{attribute 'linkalways'}
{attribute 'no_explicit_call' := 'Use the methods of this class'}
{attribute 'enable_dynamic_creation'}
FUNCTION_BLOCK DiffDrive IMPLEMENTS I_DifferentialDrive
VAR
	leftAxis : I_DriveAxis;
	rightAxis : I_DriveAxis;
	kinematics : DiffDriveKinematics;
END_VAR

METHOD Connect
VAR_INPUT
	left : I_DriveAxis;
	right : I_DriveAxis;
END_VAR
leftAxis := left;
rightAxis := right;
END_METHOD

METHOD Execute
IF leftAxis = 0 OR rightAxis = 0 THEN
	RETURN;
END_IF
leftAxis.Execute();
rightAxis.Execute();
END_METHOD

METHOD Enable
IF leftAxis = 0 OR rightAxis = 0 THEN
	RETURN;
END_IF
leftAxis.Enable();
rightAxis.Enable();
END_METHOD

METHOD Disable
IF leftAxis = 0 OR rightAxis = 0 THEN
	RETURN;
END_IF
leftAxis.Disable();
rightAxis.Disable();
END_METHOD

METHOD SetTwist
VAR_INPUT
	desiredTwist : Twist;
END_VAR
VAR
	speeds : WheelSpeeds;
END_VAR
IF leftAxis = 0 OR rightAxis = 0 THEN
	RETURN;
END_IF
speeds := kinematics.ToWheelSpeeds(desiredTwist);
leftAxis.SetVelocity(speeds.leftInMPerS);
rightAxis.SetVelocity(speeds.rightInMPerS);
END_METHOD

PROPERTY LeftWheelPositionInM : LREAL
GET
IF leftAxis <> 0 THEN
	LeftWheelPositionInM := leftAxis.PositionInM;
END_IF
END_GET
END_PROPERTY

PROPERTY RightWheelPositionInM : LREAL
GET
IF rightAxis <> 0 THEN
	RightWheelPositionInM := rightAxis.PositionInM;
END_IF
END_GET
END_PROPERTY

PROPERTY IsReady : BOOL
GET
IsReady := leftAxis <> 0 AND_THEN rightAxis <> 0 AND_THEN leftAxis.IsReady AND_THEN rightAxis.IsReady;
END_GET
END_PROPERTY

END_FUNCTION_BLOCK

(* stored: Version 1.1.0.1, ProductVersion 3.1.4026.12
   POU DiffDrive: Id {0bbf6c55-3be5-53ce-af2a-579f36f57573}, SpecialFunc None
   Method Connect: Id {097fee2a-ff23-58d4-b286-94e459e4269d}
   Method Execute: Id {faac4bfe-0ce8-591b-9cf4-3ce387f54fd0}
   Method Enable: Id {baa38bb0-278d-5e8a-871b-b137239c7090}
   Method Disable: Id {486dcacc-469b-5018-a8d0-ca66e8aaca6a}
   Method SetTwist: Id {098b0635-eb47-5c17-a9bd-67e37e18d5a2}
   Property LeftWheelPositionInM: Id {bb529295-4fcf-568d-9617-282c57c2850a}
   Get Get: Id {2965df9d-c0ea-5ec0-abec-70f400e386ad}
   Property RightWheelPositionInM: Id {e5a0aef1-afa7-5090-b787-bb6d4bf4debe}
   Get Get: Id {063c88d4-001f-54bc-8702-a0373d496641}
   Property IsReady: Id {0716dda0-318f-5c0b-9d2e-d407e343a688}
   Get Get: Id {e8c996d9-55ee-583b-8f0d-bcac8b430915} *)
